Fanuc KAREL source: kb00114.KL

-- PROVISIONAL review KL for V1013-1; original PC SHA256 80664a2ec0f5f53e5cf39ffd9108de2fc1b4f1ff760aa67e4d656856fbca2dc0
-- Incomplete behavior may be omitted. Consult companion uncertainty JSON. Do not deploy.
PROGRAM KB00114
%NOLOCKGROUP
BEGIN
  -- UNRESOLVED_PC offsets 5-14; opcodes 3F,75
  -- UNRESOLVED_PC offsets 19-26; opcodes 9D,23
  -- UNRESOLVED_PC offsets 31-49; opcodes 27,22,2A,22,31
  -- UNRESOLVED_PC offsets 54-58; opcodes 7F
END KB00114
